// Replays a CSV trajectory buffer (GVL_CsvProfile.stCsv) at the task rate. Each
// cycle it advances elapsed time, linearly interpolates BOTH channels at the same
// time index, and applies them -> the Mentee and the selected Beckhoff load motor
// stay synchronized (one player, one clock). Values are ABSOLUTE (no anchoring).
//
//   Mentee:   emits fMenteeOut; PRG_Motion routes it into the selected stCmd field
//             (setpoint_position | impedance_p_des | setpoint_velocity | setpoint_current).
//   Beckhoff: TORQUE   -> emits fLoadOut; PRG_Motion writes it to the selected
//                         motor's fTargetTorque (FB_TorqueControl streams it; the app
//                         must already be in torque mode).
//             POS/VEL  -> feeds the selected NC axis via external setpoint generation
//                         (MC_ExtSetPointGen*); the motor must be ENABLED/READY and not
//                         executing a move. VELOCITY integrates to position from the
//                         axis position captured at start.
//
// The scalar config is latched on the bStart edge; the sample arrays are read live
// (the app uploads them fully before pulsing bStart, and doesn't change them mid-run).
FUNCTION_BLOCK FB_CsvPlayer
VAR_IN_OUT
    stCsv           : ST_CsvProfile;
    AxisLoad1       : AXIS_REF;
    AxisLoad2       : AXIS_REF;
END_VAR
VAR_INPUT
    fLoad1Pos       : LREAL;    // Axis1.NcToPlc.ActPos [deg]
    fLoad2Pos       : LREAL;    // Axis2.NcToPlc.ActPos [deg]
    fDt             : REAL;     // task cycle time [s]
END_VAR
VAR_OUTPUT
    bRunning        : BOOL;
    fMenteeOut      : REAL;     // routed by PRG into the mentee field (while bRunning + enabled)
    fLoadOut        : REAL;     // routed by PRG into fTargetTorque (TORQUE domain, while bRunning + enabled)
END_VAR
VAR
    rStart          : R_TRIG;
    rStop           : R_TRIG;
    eState          : INT;
    fElapsed        : REAL;     // time into the current pass [s]
    fIdxR           : LREAL;    // fractional sample index
    iIdx            : DINT;
    fFrac           : REAL;
    fMenteeRaw      : REAL;
    fLoadRaw        : REAL;
    bWasActive      : BOOL;
    nRepDone        : UDINT;
    fRest           : REAL;

    // latched scalar config (read by the body; arrays read live from stCsv)
    nCountL         : UDINT;
    nLastIdx        : DINT;     // nCount-1
    fSampleDtL      : REAL;
    bMenteeEnL      : BOOL;
    nMenteeFieldL   : BYTE;
    bLoadEnL        : BOOL;
    nLoadMotorL     : BYTE;
    nLoadDomainL    : BYTE;
    bRepetitiveL    : BOOL;
    nRepsL          : UDINT;
    fRestSL         : REAL;

    // external setpoint generation (POSITION / VELOCITY) — instances per axis,
    // only the selected one is ever Execute'd.
    fbExt1On        : MC_ExtSetPointGenEnable;
    fbExt2On        : MC_ExtSetPointGenEnable;
    fbExt1Off       : MC_ExtSetPointGenDisable;
    fbExt2Off       : MC_ExtSetPointGenDisable;
    fbSync1         : MC_SetPosition;   // set := actual before engaging (F324/F321 guard)
    fbSync2         : MC_SetPosition;
    bSyncExec       : BOOL;     // latch: set-position sync requested / running
    bEnableExec     : BOOL;     // latch: ext-generator enable requested / running
    bSyncDone       : BOOL;
    bWaitStill      : BOOL;     // latch: waiting for NC standstill before the sync
    tonStill        : TON;      // standstill-wait timeout (proceed anyway)
    rFeedOn         : R_TRIG;   // first feed cycle -> re-anchor at engagement
    fActVelSel      : LREAL;    // selected load axis NC velocity [deg/s]
    rExtOn          : R_TRIG;
    fExtOff         : F_TRIG;
    bExtWant        : BOOL;
    bExtEnabled     : BOOL;
    fLoadStartPos   : LREAL;    // axis pos captured at start (VELOCITY integral base)
    fLoadPosAccum   : LREAL;    // VELOCITY: integral of velocity [deg]
    fExtPos         : LREAL;
    fExtVel         : LREAL;
    fPrevExtPos     : LREAL;
    nExtDir         : DINT;
END_VAR
VAR CONSTANT
    F_STILL_VELO    : LREAL := 1.0;    // NC standstill threshold [deg/s] before engaging
    T_STILL_TIMEOUT : TIME := T#2S;    // give up waiting for standstill -> proceed anyway
    ST_IDLE         : INT := 0;
    ST_RUN          : INT := 1;
    ST_REST         : INT := 2;
    ST_DONE         : INT := 3;
    DOM_TORQUE      : BYTE := 0;
    DOM_POSITION    : BYTE := 1;
    DOM_VELOCITY    : BYTE := 2;
END_VAR

rStart(CLK := stCsv.bStart);
rStop (CLK := stCsv.bStop);

IF rStop.Q THEN
    eState := ST_IDLE;
END_IF

// Start -> latch the scalar config; arrays are read live from stCsv.
IF rStart.Q AND (stCsv.nCount > 0) AND (stCsv.fSampleDt > 0.0) THEN
    nCountL       := stCsv.nCount;
    nLastIdx      := UDINT_TO_DINT(stCsv.nCount) - 1;
    fSampleDtL    := stCsv.fSampleDt;
    bMenteeEnL    := stCsv.bMenteeEnable;
    nMenteeFieldL := stCsv.nMenteeField;
    bLoadEnL      := stCsv.bLoadEnable;
    nLoadMotorL   := stCsv.nLoadMotor;
    nLoadDomainL  := stCsv.nLoadDomain;
    bRepetitiveL  := stCsv.bRepetitive;
    nRepsL        := stCsv.nReps;
    fRestSL       := stCsv.fRestS;
    fElapsed      := 0.0;
    nRepDone      := 0;
    fLoadPosAccum := 0.0;
    IF nLoadMotorL = 1 THEN fLoadStartPos := fLoad1Pos; ELSE fLoadStartPos := fLoad2Pos; END_IF
    fPrevExtPos   := fLoadStartPos;
    eState        := ST_RUN;
END_IF

bWasActive := (eState = ST_RUN) OR (eState = ST_REST);

CASE eState OF

ST_RUN:
    fIdxR := fElapsed / fSampleDtL;
    iIdx  := LREAL_TO_DINT(fIdxR);          // floor (fElapsed >= 0)
    IF iIdx >= nLastIdx THEN
        // reached the end of the table -> hold the last sample, then rep / done
        fMenteeRaw := stCsv.aMentee[nLastIdx];
        fLoadRaw   := stCsv.aLoad[nLastIdx];
        IF nLoadDomainL = DOM_VELOCITY THEN
            fLoadPosAccum := fLoadPosAccum + fLoadRaw * fDt;   // include the final sample
        END_IF
        IF NOT bRepetitiveL THEN
            eState := ST_DONE;
        ELSE
            nRepDone := nRepDone + 1;
            IF (nRepsL > 0) AND (nRepDone >= nRepsL) THEN
                eState := ST_DONE;
            ELSE
                fRest  := fRestSL;
                eState := ST_REST;
            END_IF
        END_IF
    ELSE
        fFrac      := LREAL_TO_REAL(fIdxR - DINT_TO_LREAL(iIdx));
        fMenteeRaw := stCsv.aMentee[iIdx] + fFrac * (stCsv.aMentee[iIdx + 1] - stCsv.aMentee[iIdx]);
        fLoadRaw   := stCsv.aLoad[iIdx]   + fFrac * (stCsv.aLoad[iIdx + 1]   - stCsv.aLoad[iIdx]);
        IF nLoadDomainL = DOM_VELOCITY THEN
            fLoadPosAccum := fLoadPosAccum + fLoadRaw * fDt;     // integrate velocity -> position
        END_IF
        fElapsed := fElapsed + fDt;
    END_IF

ST_REST:
    fRest := fRest - fDt;                   // hold last sample during the rest
    IF fRest <= 0.0 THEN
        fElapsed := 0.0;
        IF nLoadDomainL = DOM_VELOCITY THEN     // re-anchor so rest-drift doesn't compound
            fLoadStartPos := SEL(nLoadMotorL = 1, fLoad2Pos, fLoad1Pos);
            fLoadPosAccum := 0.0;
        END_IF
        eState := ST_RUN;
    END_IF

ST_DONE:
    ;                                       // hold last values

ST_IDLE:
    ;                                       // not running

END_CASE

//----------------------------------------------------------------------
// BECKHOFF external setpoint generation (POSITION / VELOCITY domains only).
//----------------------------------------------------------------------
bExtWant := bLoadEnL
            AND ((nLoadDomainL = DOM_POSITION) OR (nLoadDomainL = DOM_VELOCITY))
            AND ((eState = ST_RUN) OR (eState = ST_REST));
rExtOn(CLK := bExtWant);
fExtOff(CLK := bExtWant);

// Engagement chain: scrub mailbox -> wait-standstill -> sync -> enable ->
// re-anchor. See FB_LoadMotorProfile for the full F324 root-cause note:
// the PlcToNc ExtSetPos/Velo/Direction image persists between runs and the
// NC consumes it at generator activation before the first PLC feed; the
// Direction-0 scrub while engagement is pending closes that window.
IF rExtOn.Q THEN
    bWaitStill  := TRUE;                // stage 0: let the shaft settle first
    bSyncExec   := FALSE;
    bEnableExec := FALSE;
    tonStill(IN := FALSE);
END_IF
IF fExtOff.Q THEN                       // run ended/stopped mid-sequence
    bWaitStill  := FALSE;
    bSyncExec   := FALSE;
    bEnableExec := FALSE;
    tonStill(IN := FALSE);
    // disarm the mailbox: leave the last commanded position with vel 0 and
    // Direction 0, so a later engagement can never replay this run's sample
    IF nLoadMotorL = 1 THEN
        MC_ExtSetPointGenFeed(Position := fPrevExtPos, Velocity := 0.0,
                              Acceleration := 0.0, Direction := 0, Axis := AxisLoad1);
    ELSE
        MC_ExtSetPointGenFeed(Position := fPrevExtPos, Velocity := 0.0,
                              Acceleration := 0.0, Direction := 0, Axis := AxisLoad2);
    END_IF
END_IF

// stage 0: wait for NC standstill. After a high-amplitude TORQUE run the shaft
// is still creeping when the next profile starts; syncing/engaging on a moving
// shaft leaves the anchor stale by the time the first feed lands (F324).
// Timeout proceeds anyway so a slowly-drifting axis can't block the run.
IF bWaitStill THEN
    fActVelSel := SEL(nLoadMotorL = 1, AxisLoad2.NcToPlc.ActVelo, AxisLoad1.NcToPlc.ActVelo);
    tonStill(IN := TRUE, PT := T_STILL_TIMEOUT);
    IF (ABS(fActVelSel) <= F_STILL_VELO) OR tonStill.Q THEN
        tonStill(IN := FALSE);
        bWaitStill := FALSE;
        bSyncExec  := TRUE;
    END_IF
END_IF
fbSync1(Axis := AxisLoad1, Execute := bSyncExec AND (nLoadMotorL = 1),
        Position := fLoad1Pos, Mode := FALSE);
fbSync2(Axis := AxisLoad2, Execute := bSyncExec AND (nLoadMotorL = 2),
        Position := fLoad2Pos, Mode := FALSE);
bSyncDone := SEL(nLoadMotorL = 1,
                 fbSync2.Done OR fbSync2.Error,
                 fbSync1.Done OR fbSync1.Error);
IF bSyncExec AND bSyncDone THEN
    bSyncExec := FALSE;
    IF bExtWant THEN
        bEnableExec := TRUE;            // sync done -> now engage the generator
    END_IF
END_IF

fbExt1On(Axis := AxisLoad1, Execute := bEnableExec AND (nLoadMotorL = 1),
         Position := fLoad1Pos, PositionType := POSITIONTYPE_ABSOLUTE);
fbExt2On(Axis := AxisLoad2, Execute := bEnableExec AND (nLoadMotorL = 2),
         Position := fLoad2Pos, PositionType := POSITIONTYPE_ABSOLUTE);
bExtEnabled := SEL(nLoadMotorL = 1, fbExt2On.Enabled, fbExt1On.Enabled);  // selected axis
IF bEnableExec AND bExtEnabled THEN
    bEnableExec := FALSE;               // one-shot: drop Execute once engaged
END_IF

// stage 3: re-anchor at the ACTUAL engagement instant. The start-edge anchor
// is stale by the standstill-wait + sync + enable cycles; on a shaft that
// crept meanwhile the first VELOCITY command would step by that drift (F324).
// POSITION feeds absolute table values, so only the feed-forward seed applies.
rFeedOn(CLK := bExtWant AND bExtEnabled);
IF rFeedOn.Q THEN
    IF nLoadDomainL = DOM_VELOCITY THEN
        fLoadStartPos := SEL(nLoadMotorL = 1, fLoad2Pos, fLoad1Pos);
        fLoadPosAccum := 0.0;
    END_IF
    fPrevExtPos := SEL(nLoadMotorL = 1, fLoad2Pos, fLoad1Pos);
END_IF

IF bExtWant AND bExtEnabled THEN
    IF nLoadDomainL = DOM_POSITION THEN
        fExtPos := fLoadRaw;                                  // absolute position [deg]
        fExtVel := (fExtPos - fPrevExtPos) / MAX(fDt, 1E-6);  // numeric feed-forward
    ELSE
        fExtPos := fLoadStartPos + fLoadPosAccum;             // VELOCITY: start + integral
        IF eState = ST_RUN THEN fExtVel := fLoadRaw; ELSE fExtVel := 0.0; END_IF
    END_IF
    fPrevExtPos := fExtPos;

    IF   fExtVel > 0.0 THEN nExtDir := 1;
    ELSIF fExtVel < 0.0 THEN nExtDir := -1;
    ELSE                    nExtDir := 0;
    END_IF

    IF nLoadMotorL = 1 THEN
        MC_ExtSetPointGenFeed(Position := fExtPos, Velocity := fExtVel,
                              Acceleration := 0.0, Direction := nExtDir, Axis := AxisLoad1);
    ELSE
        MC_ExtSetPointGenFeed(Position := fExtPos, Velocity := fExtVel,
                              Acceleration := 0.0, Direction := nExtDir, Axis := AxisLoad2);
    END_IF
ELSIF bExtWant THEN
    // engagement pending (standstill wait / sync / enable in flight): scrub
    // the mailbox every cycle so the NC's activation window can only ever
    // see (current actual position, vel 0, Direction 0 = do not apply)
    IF nLoadMotorL = 1 THEN
        MC_ExtSetPointGenFeed(Position := fLoad1Pos, Velocity := 0.0,
                              Acceleration := 0.0, Direction := 0, Axis := AxisLoad1);
    ELSE
        MC_ExtSetPointGenFeed(Position := fLoad2Pos, Velocity := 0.0,
                              Acceleration := 0.0, Direction := 0, Axis := AxisLoad2);
    END_IF
    fPrevExtPos := SEL(nLoadMotorL = 1, fLoad2Pos, fLoad1Pos);
ELSE
    fPrevExtPos := SEL(nLoadMotorL = 1, fLoad2Pos, fLoad1Pos);   // keep the FF seed fresh
END_IF

fbExt1Off(Axis := AxisLoad1, Execute := fExtOff.Q AND (nLoadMotorL = 1));
fbExt2Off(Axis := AxisLoad2, Execute := fExtOff.Q AND (nLoadMotorL = 2));

//----------------------------------------------------------------------
// OUTPUTS / STATUS
//----------------------------------------------------------------------
fMenteeOut           := fMenteeRaw;
fLoadOut             := fLoadRaw;
bRunning             := bWasActive;
stCsv.bRunning       := bRunning;
stCsv.fElapsed       := fElapsed;
stCsv.fMenteeOut     := fMenteeRaw;
stCsv.fLoadOut       := fLoadRaw;
stCsv.bLoadExtActive := bExtWant AND bExtEnabled;

END_FUNCTION_BLOCK

(* stored: Version 1.1.0.1, ProductVersion 3.1.4026.18
   POU FB_CsvPlayer: Id {5d3b8e16-7c41-4a90-b2e7-6f1a9c3d2b58}, SpecialFunc None *)
